TYPE ST_VisuFinger :
STRUCT
	(* One gripper finger, always drawn as a cylinder. Its frame's origin is the centre of its top face; it extends
	   along its local -Z. The grip point, where a carried product's top touches, is the centre of its bottom face. *)
	fDiameter : LREAL; // mm
	fHeight : LREAL; // mm
	(* Where the finger's frame lies on the gripper flange (protocol 20, ADR 0018): position in the flange frame and
	   rotation about its Z. Clients place the finger by it while its state reports no pose (bPoseReported). *)
	stOffset : ST_VisuPlanarPose; // mm, degrees
END_STRUCT
END_TYPE

(* stored: Version 1.1.0.1, ProductVersion 3.1.4026.18
   DUT ST_VisuFinger: Id {105d6c3c-073d-47d8-b0c6-24cc6269dbd4} *)
